// TIA Portal V21 export
// export: Created 2026-11-10T07:35:27.1807692Z, ExportSetting WithDefaults, DisplayName Totally Integrated Automation Portal, DisplayVersion V21 Update 3, DisplayName STEP 7 Professional, DisplayVersion V21 Update 3, DisplayName STEP 7 Safety, DisplayVersion V21, DisplayName Tech WebApplication, DisplayVersion V21, DisplayName WinCC Basic/Comfort/Advanced, DisplayVersion V21 Update 3, DisplayName WinCC Unified, DisplayVersion V21 Update 3
FUNCTION_BLOCK "FB_Lad_ou017"   // FB83, LAD
{ S7_Optimized_Access := 'TRUE' }
VERSION : 0.1
// stored: AutoNumber true, IsIECCheckEnabled false, IsRetainMemResEnabled false, MemoryReserve 100, SetENOAutomatically false, UDAEnableTagReadback false
   VAR_INPUT
      v_req : Bool;
      v_id : CONN_OUC;
      v_len : UDInt;
   END_VAR
   VAR_OUTPUT
      v_done : Bool;
      v_busy : Bool;
      v_error : Bool;
      v_status : Word;
   END_VAR
   VAR_IN_OUT
      v_data : Array[0..99] of Byte;
      v_addr : Array[0..99] of Byte;
   END_VAR
   VAR
      inst { S7_SetPoint := 'True'} : TUSEND;
   END_VAR
BEGIN

REGION Network 1: TUSEND - Sending data
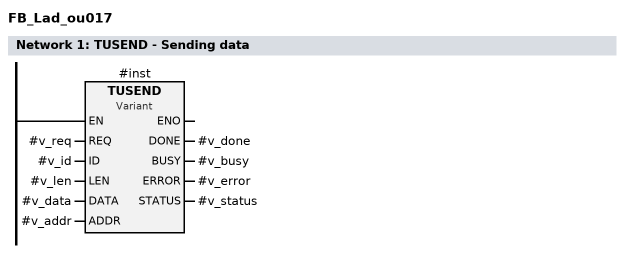
   RUNG wire#powerrail
      { S7_Templates := "[ptr_type := Variant, value_type := UDInt, id_type := CONN_OUC, addr_type := Variant]" } #inst.TUSEND(REQ := #v_req, ID := #v_id, LEN := #v_len, DONE => #v_done, BUSY => #v_busy, ERROR => #v_error, STATUS => #v_status, DATA := #v_data, ADDR := #v_addr)
   END_RUNG
   // the same network as SCL:
   #inst(REQ := #v_req,   // TUSEND
         ID := #v_id,
         LEN := #v_len,
         DATA := #v_data,
         ADDR := #v_addr,
         DONE => #v_done,
         BUSY => #v_busy,
         ERROR => #v_error,
         STATUS => #v_status);
END_REGION
END_FUNCTION_BLOCK
